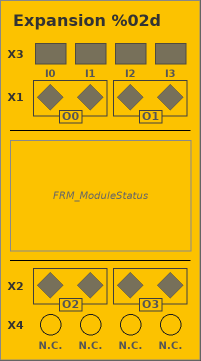
VISUALIZATION FRM_Module4DI4DOR  // 201x361
VAR_IN_OUT
    stModuleData: ST_PNOZModuleData;
END_VAR
VAR_INPUT
    nIndex: USINT;
END_VAR
    Rectangle (0,0 201x361)
    Line (10,130) (190,130)
    Line (10,260) (190,260)
    Label (0,44 31x21), "X3"
    Label (0,87 31x21), "X1"
    Label (0,276 31x21), "X2"
    Label (0,315 31x21), "X4"
    Frame (10,140 181x111)
        shows FRM_ModuleStatus(bPower := stModuleData.stLEDState.bPower, bRun := stModuleData.stLEDState.bRun, bDiag := stModuleData.stLEDState.bDiag, bFault := stModuleData.stLEDState.bFault, bInputFault := stModuleData.stLEDState.bInputFault, bOutputFault := stModuleData.stLEDState.bOutputFault, sName := stModuleData.sName, nID := stModuleData.nID, nSerialNumber := stModuleData.nSerialNumber, anRevision := stModuleData.anDeviceVersion)
    Textfield (10,0 181x41), "Expansion %02d", text variable: nIndex
    Label (30,68 41x11), "I0"
    Label (70,68 41x11), "I1"
    Label (110,68 41x11), "I2"
    Label (150,68 41x11), "I3"
    Rectangle (35,43 31x21), colour toggle: stModuleData.anInput[1].b0
    Rectangle (75,43 31x21), colour toggle: stModuleData.anInput[1].b1
    Rectangle (115,43 31x21), colour toggle: stModuleData.anInput[1].b2
    Rectangle (155,43 31x21), colour toggle: stModuleData.anInput[1].b3
    Label (30,340 41x11), "N.C."
    Label (70,340 41x11), "N.C."
    Label (110,340 41x11), "N.C."
    Label (150,340 41x11), "N.C."
    Ellipse (40,314 21x21)
    Ellipse (80,314 21x21)
    Polygon (37,285) (50,272) (63,285) (50,298) (50,298), colour toggle: stModuleData.anOutput[1].b2
    Polygon (77,285) (90,272) (103,285) (90,298) (90,298), colour toggle: stModuleData.anOutput[1].b2
    Polygon (117,285) (130,272) (143,285) (130,298) (130,298), colour toggle: stModuleData.anOutput[1].b3
    Polygon (157,285) (170,272) (183,285) (170,298) (170,298), colour toggle: stModuleData.anOutput[1].b3
    Polygon (37,97) (50,84) (63,97) (50,110) (50,110), colour toggle: stModuleData.anOutput[1].b0
    Polygon (77,97) (90,84) (103,97) (90,110) (90,110), colour toggle: stModuleData.anOutput[1].b0
    Polygon (117,97) (130,84) (143,97) (130,110) (130,110), colour toggle: stModuleData.anOutput[1].b1
    Polygon (157,97) (170,84) (183,97) (170,110) (170,110), colour toggle: stModuleData.anOutput[1].b1
    Ellipse (120,314 21x21)
    Ellipse (160,314 21x21)
    RoundedRectangle (33,80 74x36)
    RoundedRectangle (113,80 74x36)
    RoundedRectangle (33,268 74x36)
    RoundedRectangle (113,268 74x36)
    Rectangle (59,110 23x13), "O0"
    Rectangle (139,110 23x13), "O1"
    Rectangle (59,298 23x13), "O2"
    Rectangle (139,298 23x13), "O3"
END_VISUALIZATION

(* stored: Version 1.1.0.1
   Visu FRM_Module4DI4DOR: Id {8d211ab0-b6d1-070c-33ba-4a807ec23d14} *)
